// TwinCAT 3 PLC project MotionCtrl_trial1
// ProgramVersion: 3.1.4023.0
// libraries:
//   Tc2_MC2, * (Beckhoff Automation GmbH)
//   Tc2_NC, * (Beckhoff Automation GmbH)
//   Tc2_Standard, * (Beckhoff Automation GmbH)
//   Tc2_System, * (Beckhoff Automation GmbH)
//   Tc3_Module, * (Beckhoff Automation GmbH)
// project tree:
//   / PlcTask.TcTTO
//   POUs/ MAIN.TcPOU
// real-time tasks:
//   TASK PlcTask: cycle T#10ms, priority 20, ADS port 350
// motion (NC):
//   TASK NC-Task 1 SAF: cycle T#2ms, priority 4, ADS port 501
//   TASK NC-Task 1 SVB: cycle T#10ms, priority 8, ADS port 511
//   AXIS Axis 1 (id 1)
//     OtherSettings: AllowMotionCmdToSlave=true
//     encoder EncType=19
//       EncPara: MaxCount=#xffffffff
//     drive DrvType=16
//       DrvPara: MaxCount=#xffffffff, DriveControlDWord=#x00020000
//         Analog: TorqueSetpointScale=10, ScaleFactorActTorque=0.1
//         TimeComp: TaskDelayCycles=1
//     controller CtrType=1
//       CtrPara: PriorControlFactor=1
//         PosDiffControl: Enable=false
//         Observer: BandWidth=20
//   AXIS Axis 2 (id 2)
//     OtherSettings: AllowMotionCmdToSlave=true
//     encoder EncType=19
//       EncPara: MaxCount=#xffffffff
//     drive DrvType=16
//       DrvPara: MaxCount=#xffffffff, DriveControlDWord=#x00020000
//         Analog: TorqueSetpointScale=10, ScaleFactorActTorque=0.1
//         TimeComp: TaskDelayCycles=1
//     controller CtrType=1
//       CtrPara: PriorControlFactor=1
//         PosDiffControl: Enable=false
//         Observer: BandWidth=20
//   AXIS Axis 3 (id 3)
//     OtherSettings: AllowMotionCmdToSlave=true
//     encoder EncType=19
//       EncPara: MaxCount=#xffffffff
//     drive DrvType=16
//       DrvPara: MaxCount=#xffffffff, DriveControlDWord=#x00020000
//         Analog: TorqueSetpointScale=10, ScaleFactorActTorque=0.1
//         TimeComp: TaskDelayCycles=1
//     controller CtrType=1
//       CtrPara: PriorControlFactor=1
//         PosDiffControl: Enable=false
//         Observer: BandWidth=20
//   AXIS Axis 4 (id 4)
//     OtherSettings: AllowMotionCmdToSlave=true
//     encoder EncType=19
//       EncPara: MaxCount=#xffffffff
//     drive DrvType=16
//       DrvPara: MaxCount=#xffffffff, DriveControlDWord=#x00020000
//         Analog: TorqueSetpointScale=10, ScaleFactorActTorque=0.1
//         TimeComp: TaskDelayCycles=1
//     controller CtrType=1
//       CtrPara: PriorControlFactor=1
//         PosDiffControl: Enable=false
//         Observer: BandWidth=20
// I/O:
//   DEVICE Device 2 (EtherCAT), AmsNetId 169.254.233.249.3.1
//     Drive 1 (ASDA-A2-E CoE Drive) [Delta ASDA-A2-E EtherCAT(CoE) Drive Rev4]
//     Drive 2 (ASDA-A2-E CoE Drive) [Delta ASDA-A2-E EtherCAT(CoE) Drive Rev4]
//     Drive 3 (ASDA-A2-E CoE Drive) [Delta ASDA-A2-E EtherCAT(CoE) Drive Rev4]
//     Drive 4 (ASDA-A2-E CoE Drive) [Delta ASDA-A2-E EtherCAT(CoE) Drive Rev4]
// variable links:
//   NC-Task 1 SAF/Axes/Axis 1 <-> Device 2 (EtherCAT)/Drive 1 (ASDA-A2-E CoE Drive)
//     Drive/Inputs/In/nDcOutputTime <-> InfoData/DcOutputShift
//     Drive/Inputs/In/nState1 <-> 2nd TxPDO Mapping/Status Word
//     Drive/Inputs/In/nState2 <-> 2nd TxPDO Mapping/Status Word @bit 8
//     Drive/Inputs/In/nState4 @bit 1 <-> WcState/InputToggle
//     Drive/Inputs/In/nState4 <-> WcState/WcState
//     Drive/Outputs/Out/nCtrl1 <-> 2nd RxPDO Mapping/Control Word
//     Drive/Outputs/Out/nCtrl2 <-> 2nd RxPDO Mapping/Control Word @bit 8
//     Drive/Outputs/Out/nDataOut1 <-> 2nd RxPDO Mapping/TargetPosition
//     Enc/Inputs/In/nDataIn1 <-> 2nd TxPDO Mapping/ActualPosition
//     Enc/Inputs/In/nDcInputTime <-> InfoData/DcInputShift
//     Enc/Inputs/In/nState4 @bit 1 <-> WcState/InputToggle
//     Enc/Inputs/In/nState4 <-> WcState/WcState
//   NC-Task 1 SAF/Axes/Axis 2 <-> Device 2 (EtherCAT)/Drive 2 (ASDA-A2-E CoE Drive)
//     Drive/Inputs/In/nDcOutputTime <-> InfoData/DcOutputShift
//     Drive/Inputs/In/nState1 <-> 2nd TxPDO Mapping/Status Word
//     Drive/Inputs/In/nState2 <-> 2nd TxPDO Mapping/Status Word @bit 8
//     Drive/Inputs/In/nState4 @bit 1 <-> WcState/InputToggle
//     Drive/Inputs/In/nState4 <-> WcState/WcState
//     Drive/Outputs/Out/nCtrl1 <-> 2nd RxPDO Mapping/Control Word
//     Drive/Outputs/Out/nCtrl2 <-> 2nd RxPDO Mapping/Control Word @bit 8
//     Drive/Outputs/Out/nDataOut1 <-> 2nd RxPDO Mapping/TargetPosition
//     Enc/Inputs/In/nDataIn1 <-> 2nd TxPDO Mapping/ActualPosition
//     Enc/Inputs/In/nDcInputTime <-> InfoData/DcInputShift
//     Enc/Inputs/In/nState4 @bit 1 <-> WcState/InputToggle
//     Enc/Inputs/In/nState4 <-> WcState/WcState
//   NC-Task 1 SAF/Axes/Axis 3 <-> Device 2 (EtherCAT)/Drive 3 (ASDA-A2-E CoE Drive)
//     Drive/Inputs/In/nDcOutputTime <-> InfoData/DcOutputShift
//     Drive/Inputs/In/nState1 <-> 2nd TxPDO Mapping/Status Word
//     Drive/Inputs/In/nState2 <-> 2nd TxPDO Mapping/Status Word @bit 8
//     Drive/Inputs/In/nState4 @bit 1 <-> WcState/InputToggle
//     Drive/Inputs/In/nState4 <-> WcState/WcState
//     Drive/Outputs/Out/nCtrl1 <-> 2nd RxPDO Mapping/Control Word
//     Drive/Outputs/Out/nCtrl2 <-> 2nd RxPDO Mapping/Control Word @bit 8
//     Drive/Outputs/Out/nDataOut1 <-> 2nd RxPDO Mapping/TargetPosition
//     Enc/Inputs/In/nDataIn1 <-> 2nd TxPDO Mapping/ActualPosition
//     Enc/Inputs/In/nDcInputTime <-> InfoData/DcInputShift
//     Enc/Inputs/In/nState4 @bit 1 <-> WcState/InputToggle
//     Enc/Inputs/In/nState4 <-> WcState/WcState
//   NC-Task 1 SAF/Axes/Axis 4 <-> Device 2 (EtherCAT)/Drive 4 (ASDA-A2-E CoE Drive)
//     Drive/Inputs/In/nDcOutputTime <-> InfoData/DcOutputShift
//     Drive/Inputs/In/nState1 <-> 2nd TxPDO Mapping/Status Word
//     Drive/Inputs/In/nState2 <-> 2nd TxPDO Mapping/Status Word @bit 8
//     Drive/Inputs/In/nState4 @bit 1 <-> WcState/InputToggle
//     Drive/Inputs/In/nState4 <-> WcState/WcState
//     Drive/Outputs/Out/nCtrl1 <-> 2nd RxPDO Mapping/Control Word
//     Drive/Outputs/Out/nCtrl2 <-> 2nd RxPDO Mapping/Control Word @bit 8
//     Drive/Outputs/Out/nDataOut1 <-> 2nd RxPDO Mapping/TargetPosition
//     Enc/Inputs/In/nDataIn1 <-> 2nd TxPDO Mapping/ActualPosition
//     Enc/Inputs/In/nDcInputTime <-> InfoData/DcInputShift
//     Enc/Inputs/In/nState4 @bit 1 <-> WcState/InputToggle
//     Enc/Inputs/In/nState4 <-> WcState/WcState
//   MotionCtrl_trial1/MotionCtrl_trial1 Instance <-> NC-Task 1 SAF/Axes/Axis 1
//     PlcTask Inputs/MAIN.AxisList[1].NcToPlc <-> Outputs/ToPlc
//     PlcTask Outputs/MAIN.AxisList[1].PlcToNc <-> Inputs/FromPlc
//   MotionCtrl_trial1/MotionCtrl_trial1 Instance <-> NC-Task 1 SAF/Axes/Axis 2
//     PlcTask Inputs/MAIN.AxisList[2].NcToPlc <-> Outputs/ToPlc
//     PlcTask Outputs/MAIN.AxisList[2].PlcToNc <-> Inputs/FromPlc
//   MotionCtrl_trial1/MotionCtrl_trial1 Instance <-> NC-Task 1 SAF/Axes/Axis 3
//     PlcTask Inputs/MAIN.AxisList[3].NcToPlc <-> Outputs/ToPlc
//     PlcTask Outputs/MAIN.AxisList[3].PlcToNc <-> Inputs/FromPlc
//   MotionCtrl_trial1/MotionCtrl_trial1 Instance <-> NC-Task 1 SAF/Axes/Axis 4
//     PlcTask Inputs/MAIN.AxisList[4].NcToPlc <-> Outputs/ToPlc
//     PlcTask Outputs/MAIN.AxisList[4].PlcToNc <-> Inputs/FromPlc

CONFIGURATION MotionCtrl_trial1
    RESOURCE PLC ON TwinCAT3
        TASK PlcTask(INTERVAL := T#10ms, PRIORITY := 20);
        PROGRAM MAIN WITH PlcTask : MAIN;
    END_RESOURCE
END_CONFIGURATION

// ---- POUs/MAIN.TcPOU
PROGRAM MAIN
VAR CONSTANT	
	Axis_Count : INT := 4 ;
END_VAR
VAR
	power : BOOL;
	Index : INT := 1;
	
	AxisList : ARRAY[1..Axis_Count] OF AXIS_REF;
	
	Axis_State:  ARRAY[1..Axis_Count] OF INT;
	Axis_Power : ARRAY[1..Axis_Count] OF MC_Power;
	Axis_Reset : ARRAY[1..Axis_Count] OF MC_Reset;
	Axis_Home : ARRAY[1..Axis_Count] OF MC_Home;
	Axis_MoveAbs : ARRAY[1..Axis_Count] OF ARRAY[0..1] OF MC_MoveAbsolute;
	Axis_ErrorID : ARRAY[1..Axis_Count] OF UDINT;
	absSwitch : ARRAY[1..Axis_Count] OF INT;
	
	bHomeSwitch : ARRAY[1..Axis_Count] OF BOOL;
	startMove : ARRAY[1..Axis_Count] OF BOOL;
	homeBusy : ARRAY[1..Axis_Count] OF BOOL; // check if home function block is busy
	actPos : ARRAY[1..Axis_Count] OF LREAL; // array of actual position of each axis
	
	Axis_GoalPos : LREAL;
	
	rMoveVelocity : LREAL := 1600;//42666;
	rMoveAcceleration : LREAL := 12000;//120000;
	rMoveDecceleration : LREAL := 12000;//120000;
	rMoveJerk : LREAL := 560000;
	
	iCycleNum : DINT := 0;
END_VAR

iCycleNum := iCycleNum + 1;
FOR Index := 1 TO Axis_Count BY 1 DO
	AxisList[Index].ReadStatus();
	Axis_Power[Index](Axis:=AxisList[Index], Enable:=power, Enable_Positive:=TRUE, Enable_Negative:=TRUE);
	IF power THEN
		homeBusy[Index] := Axis_Home[Index].Busy;
		actPos[Index] := AxisList[Index].NcToPlc.ActPos;
		Axis_MoveAbs[Index][0](Axis:=AxisList[Index], Execute:=FALSE);
		Axis_MoveAbs[Index][1](Axis:=AxisList[Index], Execute:=FALSE);
		CASE Axis_State[Index] OF
			0: // Initial
				Axis_Reset[Index](Axis:=AxisList[Index], Execute := FALSE);
				absSwitch[Index] := 0;
				Axis_State[Index] := 10;
			10: // Start Drive Reset
				Axis_Reset[Index](Axis:=AxisList[Index], Execute := TRUE); 
				IF Axis_Reset[Index].Done THEN
					Axis_State[Index] := 20;
				ELSIF Axis_Reset[Index].Error THEN
					Axis_ErrorID[Index] := Axis_Reset[Index].ErrorID;
					Axis_State[Index] := 997;
				END_IF
			20: // Wait for Drive to Reset
				IF Axis_Power[Index].Status THEN
					Axis_State[Index] := 30;
				//ELSE
				//	Axis_State[Index] := 996;
				//	Axis_ErrorID[Index] := Axis_Power[Index].ErrorID;
				END_IF
			30: // Set current position / Homing
				IF bHomeSwitch[Index] THEN
					Axis_Home[Index](Axis:=AxisList[Index], HomingMode:=MC_HomingMode.MC_Direct, Position:=Axis_GoalPos, Execute:=TRUE);
					IF Axis_Home[Index].Error THEN
						Axis_State[Index] := 998;
					END_IF
					IF Axis_Home[Index].Done THEN
						Axis_Home[Index](Axis:=AxisList[Index], Execute:=FALSE);
						bHomeSwitch[Index] := FALSE;
					END_IF 
				ELSIF startMove[Index] THEN
					startMove[Index] := FALSE;
					Axis_State[Index] := 40;
				END_IF
			40: // Start Absolute Move
				IF Axis_MoveAbs[Index][absSwitch[Index]].Busy THEN
					absSwitch[Index] := (absSwitch[Index] + 1) MOD 2;
				END_IF
				Axis_MoveAbs[Index][absSwitch[Index]](Axis:=AxisList[Index], Position := Axis_GoalPos, BufferMode := MC_Aborting, Velocity := rMoveVelocity,
							Acceleration := rMoveAcceleration, Deceleration := rMoveDecceleration, Jerk := rMoveJerk, Execute := TRUE);
				IF Axis_MoveAbs[Index][absSwitch[Index]].Error THEN //Axis_MoveAbs.Done AND 
					Axis_State[Index] := 999;
				END_IF
				Axis_State[Index] := 30;
			
			999: //Error Fixing (TODO)
		END_CASE
	END_IF
END_FOR

END_PROGRAM
